FUNCTION_BLOCK FB_AlphaBetaFilter (* Migrated from IEC 61131-3 ST *)
  (* Standard: 61499-2 *)
  (* Version 1.0, 2026-11-06, st2fb *)
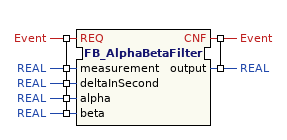
  EVENT_INPUT
    REQ WITH measurement, deltaInSecond, alpha, beta;
  END_EVENT
  EVENT_OUTPUT
    CNF WITH output;
  END_EVENT
  VAR_INPUT
    measurement : REAL;
    deltaInSecond : REAL;
    alpha : REAL;
    beta : REAL;
  END_VAR
  VAR_OUTPUT
    output : REAL;
  END_VAR
  VAR
    measurementEstimate : REAL := 0.0;
    velocityEstimate : REAL := 0.0;
    predictionError : REAL;
    measurementIntegrator : REAL;
    velocityIntegrator : REAL;
    betaResidualByDelta : REAL;
  END_VAR
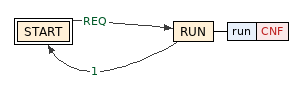
  EC_STATES
    START;
    RUN : run -> CNF;
  END_STATES
  EC_TRANSITIONS
    START TO RUN := REQ;
    RUN TO START := 1;
  END_TRANSITIONS
  ALGORITHM run IN ST:
measurementIntegrator := measurementEstimate + (velocityEstimate * deltaInSecond);
velocityIntegrator := velocityEstimate;
predictionError := measurement - measurementIntegrator;
measurementIntegrator := measurementIntegrator + (alpha * predictionError);
IF deltaInSecond > 0.0 THEN
  betaResidualByDelta := (beta * predictionError) / deltaInSecond;
ELSE
  betaResidualByDelta := 0.0;
END_IF;
velocityIntegrator := velocityIntegrator + betaResidualByDelta;
measurementEstimate := measurementIntegrator;
velocityEstimate := velocityIntegrator;
output := measurementEstimate;
  END_ALGORITHM
END_FUNCTION_BLOCK
